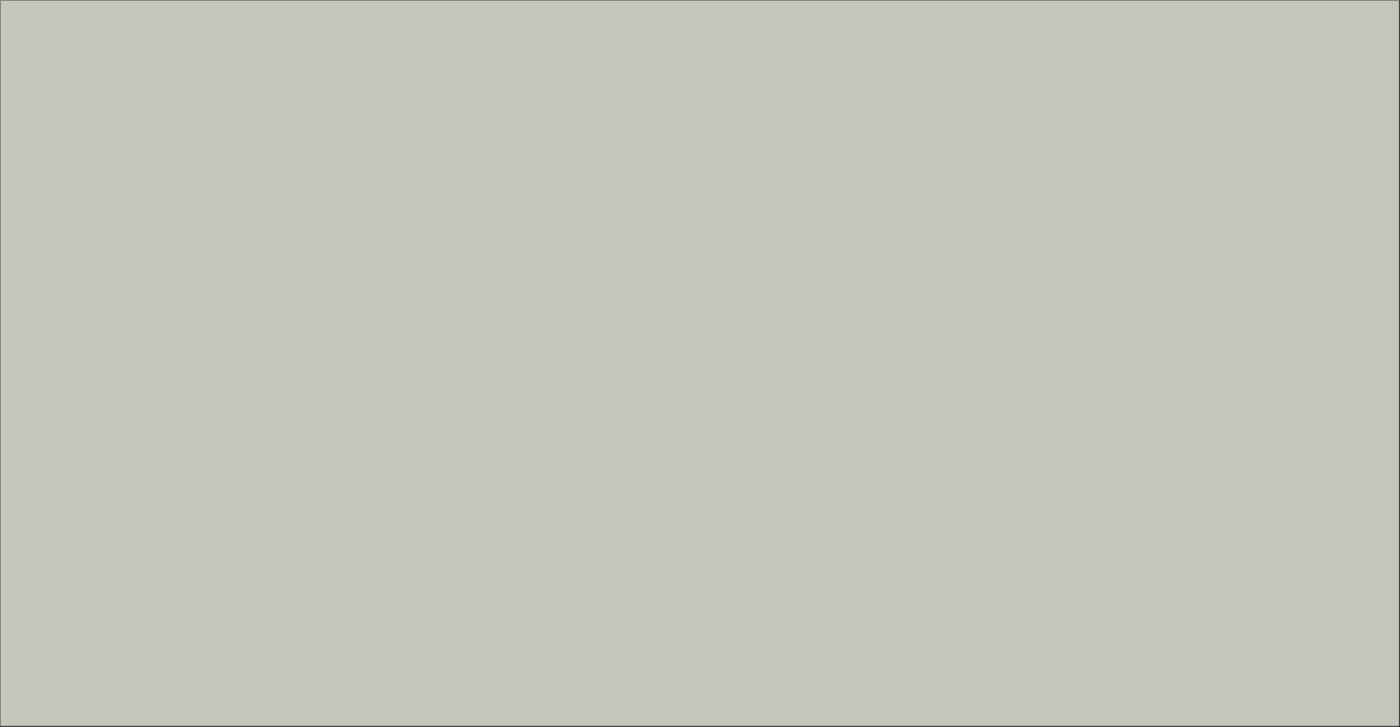
VISUALIZATION TEMP16_9_00_Content  // 1581x821
    Rectangle (0,0 1581x821)
END_VISUALIZATION

(* stored: Version 1.1.0.1, ProductVersion 3.1.4024.13
   Visu TEMP16_9_00_Content: Id {bd231165-1c89-4601-b6f4-272e29831bbb} *)
